(* IEC 61131-3 sources: llm-plc-st-eval/data/definitivo/qwen2.5-coder_14b/B7/zero_shot, 3 files *)

(* ---- ejec_1.st ---- *)
```pascal
PROGRAM SelBomba
VAR
    modoAuto : BOOL;    // Entrada que indica el modo automático
    btnManual : BOOL;   // Entrada que indica el botón manual
    nivelBajo : BOOL;  // Entrada que indica el nivel bajo
    bomba : BOOL;       // Salida que indica el estado de la bomba
END_VAR

// Lógica de selección de la fuente de mando de la bomba
IF modoAuto THEN
    // Modo automático: la bomba está encendida si nivelBajo está activo
    bomba := nivelBajo;
ELSE
    // Modo manual: la bomba obedece al botón btnManual
    bomba := btnManual;
END_IF;
```

Este programa en Structured Text (ST) cumple con los requisitos especificados. Utiliza un PROGRAM para encapsular la lógica de selección de la fuente de mando de la bomba. Las variables de entrada y salida se declaran al principio, y la lógica se implementa utilizando una estructura IF-ELSE para determinar el estado de la bomba según el modo seleccionado.

(* ---- ejec_2.st ---- *)
```pascal
PROGRAM SelBomba
VAR
    modoAuto : BOOL;  // Entrada que indica si el sistema está en modo automático
    btnManual : BOOL; // Entrada que indica el estado del botón manual
    nivelBajo : BOOL; // Entrada que indica si el nivel está por debajo del umbral
    bomba : BOOL;     // Salida que indica el estado de la bomba
END_VAR

// Lógica de selección de la fuente de mando de la bomba
IF modoAuto THEN
    // En modo automático, la bomba está encendida si nivelBajo está activo
    bomba := nivelBajo;
ELSE
    // En modo manual, la bomba obedece directamente al botón btnManual
    bomba := btnManual;
END_IF;
```

Este programa en Structured Text (ST) implementa la lógica de selección de la fuente de mando de una bomba según las especificaciones proporcionadas. La variable `bomba` indica el estado de la bomba, que depende de las entradas `modoAuto`, `btnManual` y `nivelBajo`.

(* ---- ejec_3.st ---- *)
```iec
PROGRAM SelBomba
VAR
    modoAuto : BOOL;   // Entrada que indica si el sistema está en modo automático
    btnManual : BOOL;  // Entrada que indica el estado del botón manual
    nivelBajo : BOOL;  // Entrada que indica si el nivel está por debajo del umbral
    bomba : BOOL;      // Salida que indica el estado de la bomba
END_VAR

// Lógica de selección de la fuente de mando de la bomba
IF modoAuto THEN
    // En modo automático, la bomba está encendida si nivelBajo está activo
    bomba := nivelBajo;
ELSE
    // En modo manual, la bomba obedece al botón manual
    bomba := btnManual;
END_IF;
```

Este código implementa la lógica de selección de la fuente de mando de una bomba según las especificaciones proporcionadas. La variable `bomba` indica el estado actual de la bomba basado en las entradas `modoAuto`, `btnManual` y `nivelBajo`.
